Xinje XDPPro project, PLC1: XD3-16 (software 3.8.0 2025-09-09)

PROGRAM Ladder

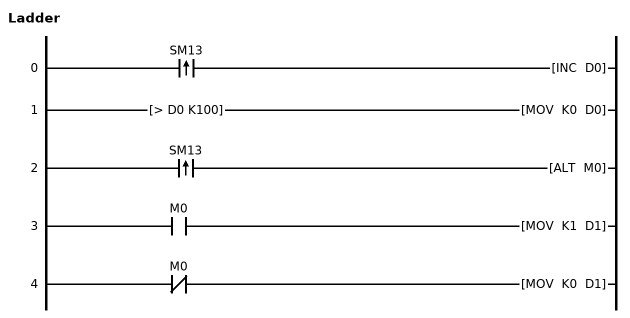
LDP    SM13
INC    D0
LD>    D0 K100
MOV    K0 D0
LDP    SM13
ALT    M0
LD     M0
MOV    K1 D1
LDI    M0
MOV    K0 D1